// TIA Portal V20 export
// export: Created 2026-10-19T18:41:55.7572766Z, ExportSetting WithDefaults, DisplayName Totally Integrated Automation Portal, DisplayVersion V20 Update 6, DisplayName TIA Portal Openness, DisplayVersion V20 Update 6, DisplayName TIA Portal Version Control Interface, DisplayVersion V20 Update 6, DisplayName SINAMICS Startdrive Advanced, DisplayVersion V20 SP1, DisplayName SINAMICS Startdrive G130, G150, S120, S150, SINAMICS MV, G220, S200, S210, DisplayVersion V20 SP1, DisplayName SINAMICS Startdrive G110M, G120, G120C, G120D, G120P, G115D, DisplayVersion V20 SP1, DisplayName STEP 7 Professional, DisplayVersion V20 Update 6, DisplayName STEP 7 Safety, DisplayVersion V20 Update 2, DisplayName WinCC Basic/Comfort/Advanced, DisplayVersion V20 Update 6, DisplayName WinCC Unified, DisplayVersion V20 Update 6
DATA_BLOCK "GateAccess_Station_FB_DB_1"   // DB425
VERSION : 0.1
// stored: AutoNumber true, DBAccessibleFromOPCUA true, InstanceOfName GateAccess_Station_FB, InstanceOfType FB
"GateAccess_Station_FB"
   // VAR_INPUT
   //    Sys_No : UInt;
   //    Right_True { ExternalAccessible := 'False'; ExternalVisible := 'False'; ExternalWritable := 'False'} : Bool;
   //    Switches { ExternalAccessible := 'False'; ExternalVisible := 'False'; ExternalWritable := 'False'} : Byte;
   //    GateLockedFeedback : Bool;
   //    NoEStop : Bool;
   //    I_G1_GuardOpen : Bool;
   //    I_L1_Unlocked : Bool;
   //    FaultResetCmd : Bool;
   //    AllDrivesHealthy : Bool;
   //    SafetyResetDone : Bool;
   //    NoVTDLocalMode : Bool;
   //    NoCrossoverPaused : Bool;
   //    Safe_Bypassed : Bool;
   //    LGX_Secure_Access : Bool;
   //    AllDevicesStopped : Bool;
   // END_VAR
   // VAR_OUTPUT
   //    Lamps { ExternalAccessible := 'False'; ExternalVisible := 'False'; ExternalWritable := 'False'} : Byte;
   //    O_S1_SolenoidEnergise : Bool;
   //    "Lock Reset" { ExternalAccessible := 'False'; ExternalVisible := 'False'; ExternalWritable := 'False'} : Bool;
   //    CurrentState : UInt;
   //    GateFault : Bool;
   // END_VAR
   // VAR_IN_OUT
   //    Gate_Station : "Gate_Station_UDT";
   // END_VAR
   // VAR
   //    RTE_PB : Bool;
   //    Reset_PB : Bool;
   //    Restart_PB : Bool;
   //    GateAccessControl : "GateAccessControl_FB";
   //    ModeManager : "ModeManager_FB";
   // END_VAR
BEGIN
END_DATA_BLOCK
